(* IEC 61131-3 sources: trust-platform/crates/trust-runtime/tests/fixtures/oscat/core/src/22_calculations, 1 file *)

(* ---- tests.st ---- *)
TEST_PROGRAM oscat_temperature_conversions_behave
ASSERT_TRUE(IN := OSCAT_BASIC_Constants());
ASSERT_NEAR(EXPECTED := REAL#77.0, ACTUAL := C_TO_F(REAL#25.0), DELTA := REAL#0.01);
ASSERT_NEAR(EXPECTED := REAL#25.0, ACTUAL := F_TO_C(REAL#77.0), DELTA := REAL#0.01);
ASSERT_NEAR(EXPECTED := REAL#298.15, ACTUAL := C_TO_K(REAL#25.0), DELTA := REAL#0.01);
ASSERT_NEAR(EXPECTED := REAL#25.0, ACTUAL := K_TO_C(REAL#298.15), DELTA := REAL#0.01);
END_TEST_PROGRAM

TEST_PROGRAM oscat_speed_and_frequency_conversions_behave
VAR
    SpeedMps : REAL;
    SpeedKmh : REAL;
    AngularFrequency : REAL;
    RoundTripFrequency : REAL;
    Period : TIME;
END_VAR

ASSERT_TRUE(IN := OSCAT_BASIC_Constants());
SpeedMps := KMH_TO_MS(REAL#36.0);
SpeedKmh := MS_TO_KMH(SpeedMps);
AngularFrequency := F_TO_OM(REAL#2.0);
RoundTripFrequency := OM_TO_F(AngularFrequency);
Period := F_TO_PT(REAL#2.0);

ASSERT_NEAR(EXPECTED := REAL#10.0, ACTUAL := SpeedMps, DELTA := REAL#0.01);
ASSERT_NEAR(EXPECTED := REAL#36.0, ACTUAL := SpeedKmh, DELTA := REAL#0.01);
ASSERT_NEAR(EXPECTED := MATH.PI2 * REAL#2.0, ACTUAL := AngularFrequency, DELTA := REAL#0.01);
ASSERT_NEAR(EXPECTED := REAL#2.0, ACTUAL := RoundTripFrequency, DELTA := REAL#0.01);
ASSERT_EQUAL(EXPECTED := INT#5, ACTUAL := MS_TO_BFT(BFT_TO_MS(INT#5)));
ASSERT_EQUAL(EXPECTED := T#500ms, ACTUAL := Period);
ASSERT_NEAR(EXPECTED := REAL#2.0, ACTUAL := PT_TO_F(T#500ms), DELTA := REAL#0.001);
END_TEST_PROGRAM

TEST_PROGRAM oscat_direction_helpers_behave
ASSERT_TRUE(IN := OSCAT_BASIC_Constants());
ASSERT_EQUAL(EXPECTED := 'N', ACTUAL := DEG_TO_DIR(INT#0, INT#1, INT#1));
ASSERT_EQUAL(EXPECTED := 'E', ACTUAL := DEG_TO_DIR(INT#90, INT#1, INT#1));
ASSERT_EQUAL(EXPECTED := 'O', ACTUAL := DEG_TO_DIR(INT#90, INT#1, INT#2));
ASSERT_EQUAL(EXPECTED := INT#90, ACTUAL := DIR_TO_DEG('E', INT#1));
ASSERT_EQUAL(EXPECTED := INT#90, ACTUAL := DIR_TO_DEG('O', INT#2));
ASSERT_EQUAL(EXPECTED := 'E', ACTUAL := LANGUAGE.DIRS[INT#1, INT#4]);
END_TEST_PROGRAM

TEST_PROGRAM oscat_geographic_conversion_behaves
ASSERT_NEAR(
    EXPECTED := REAL#59.5,
    ACTUAL := GEO_TO_DEG(INT#59, INT#30, REAL#0.0),
    DELTA := REAL#0.001
);
END_TEST_PROGRAM

TEST_FUNCTION_BLOCK oscat_energy_fb_converts_units
VAR
    Dut : ENERGY;
END_VAR

Dut(Wh := REAL#1.0);
ASSERT_NEAR(EXPECTED := REAL#3600.0, ACTUAL := Dut.YJ, DELTA := REAL#0.01);
ASSERT_NEAR(EXPECTED := REAL#1.0, ACTUAL := Dut.YWh, DELTA := REAL#0.001);
ASSERT_NEAR(EXPECTED := REAL#859.8452, ACTUAL := Dut.YC, DELTA := REAL#0.1);
END_TEST_FUNCTION_BLOCK

TEST_FUNCTION_BLOCK oscat_length_fb_converts_units
VAR
    Dut : LENGTH;
END_VAR

Dut(m := REAL#1.0);
ASSERT_NEAR(EXPECTED := REAL#1.0, ACTUAL := Dut.Ym, DELTA := REAL#0.0001);
ASSERT_NEAR(EXPECTED := REAL#39.37007874016, ACTUAL := Dut.Yin, DELTA := REAL#0.001);
ASSERT_NEAR(EXPECTED := REAL#3.28083989501, ACTUAL := Dut.Yft, DELTA := REAL#0.001);
END_TEST_FUNCTION_BLOCK

TEST_FUNCTION_BLOCK oscat_pressure_fb_converts_units
VAR
    Dut : PRESSURE;
END_VAR

Dut(bar := REAL#1.0);
ASSERT_NEAR(EXPECTED := REAL#1.0, ACTUAL := Dut.Ybar, DELTA := REAL#0.0001);
ASSERT_NEAR(EXPECTED := REAL#100000.0, ACTUAL := Dut.Ypa, DELTA := REAL#0.1);
ASSERT_NEAR(EXPECTED := REAL#0.9869232667160, ACTUAL := Dut.Yatm, DELTA := REAL#0.001);
END_TEST_FUNCTION_BLOCK

TEST_FUNCTION_BLOCK oscat_speed_fb_converts_units
VAR
    Dut : SPEED;
END_VAR

Dut(ms := REAL#10.0);
ASSERT_NEAR(EXPECTED := REAL#10.0, ACTUAL := Dut.Yms, DELTA := REAL#0.0001);
ASSERT_NEAR(EXPECTED := REAL#36.0, ACTUAL := Dut.Ykmh, DELTA := REAL#0.001);
ASSERT_NEAR(EXPECTED := REAL#22.369362920544, ACTUAL := Dut.Ymh, DELTA := REAL#0.001);
END_TEST_FUNCTION_BLOCK

TEST_FUNCTION_BLOCK oscat_temperature_fb_converts_units
VAR
    Dut : TEMPERATURE;
END_VAR

Dut(
    K := REAL#0.0,
    C := REAL#25.0,
    F := REAL#-459.67,
    Re := REAL#-218.52,
    Ra := REAL#0.0
);
ASSERT_NEAR(EXPECTED := REAL#298.15, ACTUAL := Dut.YK, DELTA := REAL#0.01);
ASSERT_NEAR(EXPECTED := REAL#25.0, ACTUAL := Dut.YC, DELTA := REAL#0.01);
ASSERT_NEAR(EXPECTED := REAL#77.0, ACTUAL := Dut.YF, DELTA := REAL#0.01);
END_TEST_FUNCTION_BLOCK

TEST_FUNCTION_BLOCK oscat_astro_fb_converts_units
VAR
    Dut : ASTRO;
END_VAR

Dut(AE := REAL#1.0);
ASSERT_NEAR(EXPECTED := REAL#149597870000.0, ACTUAL := Dut.Ym, DELTA := REAL#1000000.0);
ASSERT_NEAR(EXPECTED := REAL#1.0, ACTUAL := Dut.YAE, DELTA := REAL#0.0001);
ASSERT_NEAR(EXPECTED := REAL#4.8481322570E-6, ACTUAL := Dut.YPC, DELTA := REAL#1.0E-9);
ASSERT_NEAR(EXPECTED := REAL#1.5812776724E-5, ACTUAL := Dut.YLJ, DELTA := REAL#1.0E-8);
END_TEST_FUNCTION_BLOCK
